(* Tests F_ParseHttpUrl, which the HTTP log and span exporters use to split their endpoint URL. *)
FUNCTION_BLOCK FB_TestHttpUrlParser EXTENDS FB_TestSuite

THIS^.testHttpWithPortAndPath();
THIS^.testHttpDefaultsPortAndPath();
THIS^.testHttpsDefaultsPort();
THIS^.testRejectsMissingScheme();
THIS^.testRejectsUpperCaseScheme();
THIS^.testRejectsEmptyPort();
THIS^.testRejectsZeroPort();
THIS^.testRejectsEmptyHost();

(* An explicit port and path are split out. *)
METHOD testHttpWithPortAndPath : REFERENCE TO FB_Test
VAR
	endpoint: ST_HttpEndpoint;
END_VAR
TcUnit.TEST('testHttpWithPortAndPath');
	THIS^.AssertEquals_BOOL(TRUE, F_ParseHttpUrl(url:='http://192.168.1.10:4318/v1/traces', endpoint=>endpoint), 'Expected the URL to parse');
	THIS^.AssertEquals_BOOL(FALSE, endpoint.useTls, 'Expected plain HTTP (useTls FALSE)');
	THIS^.AssertEquals_STRING('192.168.1.10', endpoint.host, 'Expected host 192.168.1.10');
	THIS^.AssertEquals_UINT(4318, endpoint.port, 'Expected port 4318');
	THIS^.AssertEquals_STRING('/v1/traces', endpoint.path, 'Expected path /v1/traces');
TcUnit.TEST_FINISHED();
END_METHOD

(* http without a port or path uses port 80 and '/'. *)
METHOD testHttpDefaultsPortAndPath : REFERENCE TO FB_Test
VAR
	endpoint: ST_HttpEndpoint;
END_VAR
TcUnit.TEST('testHttpDefaultsPortAndPath');
	THIS^.AssertEquals_BOOL(TRUE, F_ParseHttpUrl(url:='http://collector', endpoint=>endpoint), 'Expected the URL to parse');
	THIS^.AssertEquals_BOOL(FALSE, endpoint.useTls, 'Expected plain HTTP (useTls FALSE)');
	THIS^.AssertEquals_STRING('collector', endpoint.host, 'Expected host collector');
	THIS^.AssertEquals_UINT(80, endpoint.port, 'Expected the default http port 80');
	THIS^.AssertEquals_STRING('/', endpoint.path, 'Expected the default path /');
TcUnit.TEST_FINISHED();
END_METHOD

(* https uses TLS and port 443. *)
METHOD testHttpsDefaultsPort : REFERENCE TO FB_Test
VAR
	endpoint: ST_HttpEndpoint;
END_VAR
TcUnit.TEST('testHttpsDefaultsPort');
	THIS^.AssertEquals_BOOL(TRUE, F_ParseHttpUrl(url:='https://collector/v1/logs', endpoint=>endpoint), 'Expected the URL to parse');
	THIS^.AssertEquals_BOOL(TRUE, endpoint.useTls, 'Expected HTTPS (useTls TRUE)');
	THIS^.AssertEquals_STRING('collector', endpoint.host, 'Expected host collector');
	THIS^.AssertEquals_UINT(443, endpoint.port, 'Expected the default https port 443');
	THIS^.AssertEquals_STRING('/v1/logs', endpoint.path, 'Expected path /v1/logs');
TcUnit.TEST_FINISHED();
END_METHOD

(* A URL without http:// or https:// is rejected. *)
METHOD testRejectsMissingScheme : REFERENCE TO FB_Test
VAR
	endpoint: ST_HttpEndpoint;
END_VAR
TcUnit.TEST('testRejectsMissingScheme');
	THIS^.AssertEquals_BOOL(FALSE, F_ParseHttpUrl(url:='not-a-valid-url', endpoint=>endpoint), 'Expected a URL without a scheme to be rejected');
TcUnit.TEST_FINISHED();
END_METHOD

(* The scheme must be lower case. *)
METHOD testRejectsUpperCaseScheme : REFERENCE TO FB_Test
VAR
	endpoint: ST_HttpEndpoint;
END_VAR
TcUnit.TEST('testRejectsUpperCaseScheme');
	THIS^.AssertEquals_BOOL(FALSE, F_ParseHttpUrl(url:='HTTP://collector', endpoint=>endpoint), 'Expected an upper-case scheme to be rejected');
TcUnit.TEST_FINISHED();
END_METHOD

(* A colon without a port is rejected. *)
METHOD testRejectsEmptyPort : REFERENCE TO FB_Test
VAR
	endpoint: ST_HttpEndpoint;
END_VAR
TcUnit.TEST('testRejectsEmptyPort');
	THIS^.AssertEquals_BOOL(FALSE, F_ParseHttpUrl(url:='http://collector:/v1/traces', endpoint=>endpoint), 'Expected a colon without a port to be rejected');
TcUnit.TEST_FINISHED();
END_METHOD

(* Port 0, or a port that is not a number, is rejected. *)
METHOD testRejectsZeroPort : REFERENCE TO FB_Test
VAR
	endpoint: ST_HttpEndpoint;
END_VAR
TcUnit.TEST('testRejectsZeroPort');
	THIS^.AssertEquals_BOOL(FALSE, F_ParseHttpUrl(url:='http://collector:0/v1/traces', endpoint=>endpoint), 'Expected port 0 to be rejected');
	THIS^.AssertEquals_BOOL(FALSE, F_ParseHttpUrl(url:='http://collector:abc/v1/traces', endpoint=>endpoint), 'Expected a non-numeric port to be rejected');
TcUnit.TEST_FINISHED();
END_METHOD

(* A URL without a host is rejected. *)
METHOD testRejectsEmptyHost : REFERENCE TO FB_Test
VAR
	endpoint: ST_HttpEndpoint;
END_VAR
TcUnit.TEST('testRejectsEmptyHost');
	THIS^.AssertEquals_BOOL(FALSE, F_ParseHttpUrl(url:='http:///v1/traces', endpoint=>endpoint), 'Expected a URL without a host to be rejected');
TcUnit.TEST_FINISHED();
END_METHOD

END_FUNCTION_BLOCK

(* stored: Version 1.1.0.1
   POU FB_TestHttpUrlParser: Id {fd4a6579-122f-4581-aaee-5a4ed1aab431}, SpecialFunc None
   Method testHttpWithPortAndPath: Id {36103b9b-7122-4e41-90f3-4d14ce5805c6}
   Method testHttpDefaultsPortAndPath: Id {bac255d6-5472-4ca6-bbf3-0a3b0fad9250}
   Method testHttpsDefaultsPort: Id {96033edf-ce43-4bb2-a975-a9fe09faefa0}
   Method testRejectsMissingScheme: Id {75bcad19-ec29-4de9-b9ff-0fe681a589ef}
   Method testRejectsUpperCaseScheme: Id {ddefebc6-78e3-4c5c-988f-e3eb7ba0a01d}
   Method testRejectsEmptyPort: Id {59ec2ff7-31a6-459c-bf98-4eb5e60c3267}
   Method testRejectsZeroPort: Id {45201107-0cab-4a50-b607-cef86b169fad}
   Method testRejectsEmptyHost: Id {aaf0917b-a040-42b2-bc7e-f7bff1976572} *)
